(* IEC 61131-3 sources: plcassist-cli/packages/volt-lsp-iec/test-corpus/awa-palletizer/Device/Plc Logic/Application/Library Manager/L_SUDP_SlaveUpDownloadManager, 43 files *)

(* ---- DECIMALTOHEXSTRING.fun ---- *)
FUNCTION DECIMALTOHEXSTRING : STRING
VAR_INPUT
	DWVALUE : DWORD;
	NMAXBYTESIZE : INT;
END_VAR
END_FUNCTION

(* ---- GETBOOLEANPROPERTY.fun ---- *)
FUNCTION GETBOOLEANPROPERTY : BOOL
VAR_INPUT
	STKEY : WSTRING;
END_VAR
END_FUNCTION

(* ---- GETCOMPANY.fun ---- *)
FUNCTION GETCOMPANY : WSTRING
END_FUNCTION

(* ---- GETNUMBERPROPERTY.fun ---- *)
FUNCTION GETNUMBERPROPERTY : DINT
VAR_INPUT
	STKEY : WSTRING;
END_VAR
END_FUNCTION

(* ---- GETTEXTPROPERTY.fun ---- *)
FUNCTION GETTEXTPROPERTY : WSTRING
VAR_INPUT
	STKEY : WSTRING;
END_VAR
END_FUNCTION

(* ---- GETTEXTPROPERTY2.fun ---- *)
FUNCTION GETTEXTPROPERTY2 : POINTER TO WSTRING
VAR_INPUT
	STKEY : WSTRING;
END_VAR
END_FUNCTION

(* ---- GETTITLE.fun ---- *)
FUNCTION GETTITLE : WSTRING
END_FUNCTION

(* ---- GETVERSION.fun ---- *)
FUNCTION GETVERSION : VERSION
END_FUNCTION

(* ---- GETVERSIONPROPERTY.fun ---- *)
FUNCTION GETVERSIONPROPERTY : VERSION
VAR_INPUT
	STKEY : WSTRING;
END_VAR
END_FUNCTION

(* ---- L_EXISTALLFILES.fun ---- *)
FUNCTION L_EXISTALLFILES : BOOL
END_FUNCTION

(* ---- L_PATHFIRMWAREFILES.fun ---- *)
FUNCTION L_PATHFIRMWAREFILES : STRING(L_SUDP_MAX_STRING_LENGTH.FILE_PATH)
END_FUNCTION

(* ---- L_PATHPARAMETERSETFILES.fun ---- *)
FUNCTION L_PATHPARAMETERSETFILES : STRING(L_SUDP_MAX_STRING_LENGTH.FILE_PATH)
END_FUNCTION

(* ---- L_SUDP_CRC32FINISH.fun ---- *)
FUNCTION L_SUDP_CRC32FINISH : DWORD
VAR_INPUT
	ULCRC : DWORD;
END_VAR
END_FUNCTION

(* ---- L_SUDP_CRC32INIT.fun ---- *)
FUNCTION L_SUDP_CRC32INIT : DWORD
END_FUNCTION

(* ---- L_SUDP_CRC32UPDATE.fun ---- *)
FUNCTION L_SUDP_CRC32UPDATE : DWORD
VAR_INPUT
	ULCRC : DWORD;
	PDATA : POINTER TO BYTE;
	ULSIZE : __XWORD;
END_VAR
END_FUNCTION

(* ---- L_SUDP_GETBINARYFILENAME.fun ---- *)
FUNCTION L_SUDP_GETBINARYFILENAME : BOOL
VAR_INPUT
	WFIELDBUSMASTERID : WORD;
	WINTERFACE : WORD;
	DNNODEADDRESS : DINT;
	PSBINARYFILENAME : POINTER TO STRING(20);
END_VAR
END_FUNCTION

(* ---- L_SUDP_GETBUFFERINDEX.fun ---- *)
FUNCTION L_SUDP_GETBUFFERINDEX : WORD
VAR_INPUT
	DWLENGTH : DWORD;
	DWTASKINTERVAL : DWORD;
	PERROR : POINTER TO L_SUDP_ErrorCodes;
END_VAR
END_FUNCTION

(* ---- L_SUDP_GETFBCONTROL.fun ---- *)
FUNCTION L_SUDP_GETFBCONTROL : L_SUDP_Control
VAR_INPUT
	HREGISTRATION : CAA.HANDLE;
END_VAR
END_FUNCTION

(* ---- L_SUDP_GETFWDLMODE.fun ---- *)
FUNCTION L_SUDP_GETFWDLMODE : BYTE
END_FUNCTION

(* ---- L_SUDP_GETLEMREGISTRATIONHANDLE.fun ---- *)
FUNCTION L_SUDP_GETLEMREGISTRATIONHANDLE : RTS_IEC_HANDLE
END_FUNCTION

(* ---- L_SUDP_GETPATHBOOTDIRECTORY.fun ---- *)
FUNCTION L_SUDP_GETPATHBOOTDIRECTORY : STRING(L_SUDP_MAX_STRING_LENGTH.FILE_PATH)
END_FUNCTION

(* ---- L_SUDP_GETPATHTEMPDIRECTORY.fun ---- *)
FUNCTION L_SUDP_GETPATHTEMPDIRECTORY : STRING(L_SUDP_MAX_STRING_LENGTH.FILE_PATH)
END_FUNCTION

(* ---- L_SUDP_GETPOINTERTOBUFFER.fun ---- *)
FUNCTION L_SUDP_GETPOINTERTOBUFFER : POINTER TO BYTE
VAR_INPUT
	WBUFFERNUMBER : WORD;
	PERROR : POINTER TO L_SUDP_ErrorCodes;
END_VAR
END_FUNCTION

(* ---- L_SUDP_GETTARGETVERSION.fun ---- *)
FUNCTION L_SUDP_GETTARGETVERSION : BOOL
VAR_INPUT
	ETRANSFERTYPE : L_SUDP_TransferType;
	WFIELDBUSMASTERID : WORD;
	WINTERFACE : WORD;
	DNNODEADDRESS : DINT;
	PSTARGETVERSION : POINTER TO STRING(20);
END_VAR
END_FUNCTION

(* ---- L_SUDP_ISBOOTAPPLICATIONLOADED.fun ---- *)
FUNCTION L_SUDP_ISBOOTAPPLICATIONLOADED : BOOL
END_FUNCTION

(* ---- L_SUDP_REGISTER.fun ---- *)
FUNCTION L_SUDP_REGISTER : CAA.HANDLE
VAR_INPUT
	ETRANSFERTYPE : L_SUDP_TransferType;
	WFIELDBUSMASTERID : WORD;
	WINTERFACE : WORD;
	DNNODEADDRESS : DINT;
END_VAR
END_FUNCTION

(* ---- L_SUDP_RELEASEBUFFERINDEX.fun ---- *)
FUNCTION L_SUDP_RELEASEBUFFERINDEX : BOOL
VAR_INPUT
	WBUFFERINDEX : WORD;
	PERROR : POINTER TO L_SUDP_ErrorCodes;
END_VAR
END_FUNCTION

(* ---- L_SUDP_RELEASEBUFFERINDEXWITHERROR.fun ---- *)
FUNCTION L_SUDP_RELEASEBUFFERINDEXWITHERROR : BOOL
VAR_INPUT
	WBUFFERINDEX : WORD;
	PERROR : POINTER TO L_SUDP_ErrorCodes;
END_VAR
END_FUNCTION

(* ---- L_SUDP_SENDEVENTBUSISPREOP.fun ---- *)
FUNCTION L_SUDP_SENDEVENTBUSISPREOP : BOOL
VAR_INPUT
	WFIELDBUSMASTERID : WORD;
	WINTERFACE : WORD;
END_VAR
END_FUNCTION

(* ---- L_SUDP_SETCANCONFIGURATIONDONE.fun ---- *)
FUNCTION L_SUDP_SETCANCONFIGURATIONDONE : BOOL
VAR_INPUT
	WFIELDBUSMASTERID : WORD;
	WINTERFACE : WORD;
	BYCOUNTOFSLAVE : BYTE;
END_VAR
END_FUNCTION

(* ---- L_SUDP_SETNEWFBERROR.fun ---- *)
FUNCTION L_SUDP_SETNEWFBERROR : BOOL
VAR_INPUT
	HREGISTRATION : CAA.HANDLE;
	EERROR : L_SUDP_ErrorCodes;
END_VAR
END_FUNCTION

(* ---- L_SUDP_SETNEWFBPROGRESS.fun ---- *)
FUNCTION L_SUDP_SETNEWFBPROGRESS : BOOL
VAR_INPUT
	HREGISTRATION : CAA.HANDLE;
	BYPROGRESS : BYTE;
END_VAR
END_FUNCTION

(* ---- L_SUDP_SETNEWFBSTATE.fun ---- *)
FUNCTION L_SUDP_SETNEWFBSTATE : BOOL
VAR_INPUT
	HREGISTRATION : CAA.HANDLE;
	ESTATE : L_SUDP_State;
END_VAR
END_FUNCTION

(* ---- L_SUDP_UPDOWNLOADFBEXIT.fun ---- *)
FUNCTION L_SUDP_UPDOWNLOADFBEXIT : BOOL
VAR_INPUT
	WFIELDBUSMASTERID : WORD;
	WINTERFACE : WORD;
	ETRANSFERTYPE : L_SUDP_TransferType;
END_VAR
END_FUNCTION

(* ---- L_SUDP_UPDOWNLOADFBINIT.fun ---- *)
FUNCTION L_SUDP_UPDOWNLOADFBINIT : BOOL
VAR_INPUT
	WFIELDBUSMASTERID : WORD;
	WINTERFACE : WORD;
	ETRANSFERTYPE : L_SUDP_TransferType;
END_VAR
END_FUNCTION

(* ---- L_SUDP_WRITEERRORMESSAGE.fun ---- *)
FUNCTION L_SUDP_WRITEERRORMESSAGE : BOOL
VAR_INPUT
	HLEMACCESS : RTS_IEC_HANDLE;
	SDEVICENAME : STRING;
	WSLAVEADR : WORD;
	TRANSFERTYPE : L_SUDP_TransferType;
	ERRORCODE : L_SUDP_ErrorCodes;
	PSERRORATTACHMENT : POINTER TO STRING;
END_VAR
END_FUNCTION

(* ---- L_SUDP_WRITEERRORMESSAGEWITHLOGCLASS.fun ---- *)
FUNCTION L_SUDP_WRITEERRORMESSAGEWITHLOGCLASS : BOOL
VAR_INPUT
	HLEMACCESS : RTS_IEC_HANDLE;
	SDEVICENAME : STRING;
	WSLAVEADR : WORD;
	TRANSFERTYPE : L_SUDP_TransferType;
	LOGCLASS : UDINT;
	ERRORCODE : L_SUDP_ErrorCodes;
	PSERRORATTACHMENT : POINTER TO STRING;
END_VAR
END_FUNCTION

(* ---- L_SUDP_WRITELOGMESSAGE.fun ---- *)
FUNCTION L_SUDP_WRITELOGMESSAGE : BOOL
VAR_INPUT
	HLEMACCESS : RTS_IEC_HANDLE;
	SDEVICENAME : STRING;
	WSLAVEADR : WORD;
	TRANSFERTYPE : L_SUDP_TransferType;
	LOGCLASS : UDINT;
	UDILOGID : UDINT;
	PSLOGMESSAGE : POINTER TO STRING;
END_VAR
END_FUNCTION

(* ---- L_SUDP_WRITENEWPARSETCHECKSUM.fun ---- *)
FUNCTION L_SUDP_WRITENEWPARSETCHECKSUM : BOOL
VAR_INPUT
	EBUSTYPE : L_SUDP_BUS_TYPE;
	WNETID : WORD;
	WSLAVEADR : WORD;
	DWFILECRC : DWORD;
END_VAR
END_FUNCTION

(* ---- L_SUDP_WRITESUCCESSMESSAGE.fun ---- *)
FUNCTION L_SUDP_WRITESUCCESSMESSAGE : BOOL
VAR_INPUT
	HLEMACCESS : RTS_IEC_HANDLE;
	SDEVICENAME : STRING;
	WSLAVEADR : WORD;
	TRANSFERTYPE : L_SUDP_TransferType;
	SUCCESSCODE : L_SUDP_SuccessCodes;
	PSATTACHEDTXT : POINTER TO STRING;
END_VAR
END_FUNCTION

(* ---- CALCULATECHECKSUMFROMOPENFILE.fb ---- *)
FUNCTION_BLOCK CALCULATECHECKSUMFROMOPENFILE EXTENDS AsyncBaseClass
VAR_INPUT
	XEXECUTE : BOOL;
	HPARAFILE : RTS_IEC_HANDLE;
	DWFILESIZE : __XWORD;
	PBYBUFFER : POINTER TO BYTE;
	SZBUFFERSIZE : __XWORD;
	DWFILEOFFSETCHECKSUMCALC : DWORD;
	DWPOSITIONCHECKSUM : __XWORD := 32;
END_VAR
VAR_OUTPUT
	XDONE : BOOL;
	XERROR : BOOL;
	EERROR : L_SUDP_ErrorCodes;
	ULCRC32 : UDINT;
END_VAR
VAR
	JOB : RTS_IEC_HANDLE := CAA.gc_hINVALID;
	JOBSTATE : UDINT;
	RESULTTASK : RTS_IEC_RESULT;
	ASYNCJOBPARAM : AsyncJob_Param;
	ASYNCJOBNAME : STRING := 'UploacCalcCRC';
	RESULTASYNCADD : UDINT;
	XEXECUTEOLD : BOOL;
	DWFILEPOS : __XWORD;
	A : INT;
END_VAR
END_FUNCTION_BLOCK

METHOD DOJOB : RTS_IEC_RESULT
END_METHOD

METHOD DUMMYJOB : RTS_IEC_RESULT
END_METHOD

METHOD FB_EXIT : BOOL
VAR_INPUT
	BINCOPYCODE : BOOL;
END_VAR
END_METHOD

METHOD FB_INIT : BOOL
VAR_INPUT
	BINITRETAINS : BOOL;
	BINCOPYCODE : BOOL;
END_VAR
END_METHOD

(* ---- L_SUDP_PRMFILE_READWRITE.fb ---- *)
FUNCTION_BLOCK L_SUDP_PRMFILE_READWRITE
VAR_INPUT
	XEXECUTE : BOOL;
	EBUSTYPE : L_SUDP_BUS_TYPE;
	WNETID : WORD := 0;
	WSLAVEADR : WORD := 1;
	SDEVICENAME : STRING;
	HREGISTRATION : CAA.HANDLE := CAA.gc_hINVALID;
	SFULLFILENAME : STRING(L_SUDP_MAX_STRING_LENGTH.PATH_AND_FILE_NAME);
	UDITIMEOUT : UDINT := 500000;
	DWFILEOFFSETCHECKSUMCALC : DWORD;
END_VAR
VAR_OUTPUT
	XDONE : BOOL;
	XERROR : BOOL;
	EERROR : L_SUDP_ErrorCodes;
	PSATTACHEDERRORTXT : POINTER TO STRING;
END_VAR
VAR
	STATE : L_SUDP_PRM_FILE_READWRITE_STATES := L_SUDP_PRM_FILE_READWRITE_STATES.NONE;
	XEXECUTEOLD : BOOL;
	XREPLACEOLDFILE : BOOL;
	FGETFS : FILE.GetSize;
	FOPEN : FILE.Open;
	FREAD : FILE.Read;
	FWRITE : FILE.Write;
	FCLOSE : FILE.Close;
	FSETPOS : FILE.SetPos;
	FRENAME : FILE.Rename;
	FDELETE : FILE.Delete;
	UDITIMEOUTFILEACCESS : UDINT := 200000;
	CALCCRC : CalculateChecksumFromOpenFile;
	HPARAFILEREAD : CAA.HANDLE;
	HPARAFILEWRITE : RTS_IEC_HANDLE;
	PIOBUFFER : POINTER TO BYTE;
	ADWHEADER : ARRAY [0..((((SIZEOF(L_SUDP_PAR_FILE_HDR) + SIZEOF(L_SUDP_PAR_DATA_HDR)) - 1) / SIZEOF(DWORD)) + 1)] OF DWORD;
	ADWIOBUFFER : ARRAY [0..66] OF DWORD;
	XFIRSTPARAMHEADERWASREAD : BOOL;
	ADWSDOVALUEBUFFER : ARRAY [0..66] OF DWORD;
	DWPARDATASZ : DWORD;
	DWPARDATAPOSITION : DWORD;
	DWNEWPARDATAPOSITION : DWORD;
	PFILEHDR : POINTER TO L_SUDP_PAR_FILE_HDR;
	PPARDATHDR : POINTER TO L_SUDP_PAR_DATA_HDR;
	PARAMHDR : L_SUDP_PARM_HDR;
	PPARAMHDR : POINTER TO L_SUDP_PARM_HDR;
	SZPARAFILESZ : UDINT;
	SDODATALENGTH : UINT;
	SDOVALUEREADDONE : BOOL;
	DWCRC32 : DWORD;
	DWCRC32FILEPOSITION : DWORD;
	MYTESTCOUNTER : INT;
END_VAR
END_FUNCTION_BLOCK

METHOD BEFORESTARTEXECUTION
END_METHOD

METHOD READVALUEFROMFIELDBUS_LOOP : INT
END_METHOD

METHOD READVALUEFROMFIELDBUS_START
VAR_INPUT
	PARAMHDR : POINTER TO L_SUDP_PARM_HDR;
	PBYBUFFER : POINTER TO BYTE;
	SZBUFFERSIZE : UINT;
END_VAR
END_METHOD

METHOD FB_EXIT : BOOL
VAR_INPUT
	BINCOPYCODE : BOOL;
END_VAR
END_METHOD

(* ---- L_SUDP_UPDOWNLOAD.fb ---- *)
FUNCTION_BLOCK L_SUDP_UPDOWNLOAD
VAR_OUTPUT
	ESTATE : L_SUDP_State;
	EERROR : L_SUDP_ErrorCodes;
	BYPROGRESS : BYTE;
END_VAR
VAR
	EBUSTYPE : L_SUDP_BUS_TYPE;
	WNETID : WORD;
	WSLAVEADR : WORD;
	TRANSFERTYPE : L_SUDP_TransferType;
	DWTASKINTERVAL : DWORD;
	PTASKINFO : POINTER TO CmpIecTask.Task_Info2;
	HTASKHANDLE : RTS_IEC_HANDLE;
	ETASKRESULT : RTS_IEC_RESULT;
	BFIRSTINITIALIZEDONE : BOOL;
	BREGISTERTODOWNLOADMANAGERDONE : BOOL;
	HREGISTRATION : CAA.HANDLE := CAA.gc_hINVALID;
	PBYDLUPMGRBUFFER : POINTER TO BYTE;
	WBUFFERINDEX : WORD := SINT_TO_WORD((0 - 1));
	M_HLEMACCESS : RTS_IEC_HANDLE;
	FILE_IO_TIMEOUT_FACTOR : UDINT := 10000;
	ETC_SDO_TIMEOUT_FACTOR : UDINT := 1;
	ETC_FOE_TIMEOUT_FACTOR : UDINT := 5;
	ETC_SET_STATE_TIMEOUT_FACTOR : UDINT := 5;
	PARSET_FILE_TYPE_INVALID : DWORD := 0;
	PARSET_FILE_TYPE_9400 : DWORD := 1;
	PARSET_FILE_TYPE_I700_STORE : DWORD := 2;
	PARSET_FILE_TYPE_I700_ALL : DWORD := 3;
	PARSET_FILE_TYPE_STANDARD : DWORD := 1000;
	INVALID_BUFFER_INDEX : WORD := SINT_TO_WORD((0 - 1));
	LEMACCESSHANDLE : RTS_IEC_HANDLE;
END_VAR
END_FUNCTION_BLOCK

METHOD FB_EXIT : BOOL
VAR_INPUT
	BINCOPYCODE : BOOL;
END_VAR
END_METHOD

METHOD FIRSTINITIALIZE
VAR_INPUT
	PIOCONFIGCONNECTOR : POINTER TO IoConfigConnector;
END_VAR
END_METHOD

METHOD GETPARAMETERSETFILENAME : BOOL
VAR_INPUT
	EFIELDBUSMASTERID : L_SUDP_BUS_TYPE;
	WNETID : WORD;
	WSLAVEADR : WORD;
	PPATHBUFFER : POINTER TO STRING;
END_VAR
VAR_OUTPUT
	BRETC : BOOL := TRUE;
END_VAR
END_METHOD

METHOD GETDWTASKINTERVAL
END_METHOD

METHOD REGISTERFBTODLUPMGR : BOOL
VAR_INPUT
	PIOCONFIGCONNECTOR : POINTER TO IoConfigConnector;
END_VAR
END_METHOD
